// TIA Portal V21 export
// export: Created 2026-11-10T19:21:32.9271764Z, ExportSetting WithDefaults, DisplayName Totally Integrated Automation Portal, DisplayVersion V21 Update 3, DisplayName STEP 7 Professional, DisplayVersion V21 Update 3, DisplayName STEP 7 Safety, DisplayVersion V21, DisplayName Tech WebApplication, DisplayVersion V21, DisplayName WinCC Basic/Comfort/Advanced, DisplayVersion V21 Update 3, DisplayName WinCC Unified, DisplayVersion V21 Update 3
FUNCTION_BLOCK "FB_Lad_pt007"   // FB2, LAD
{ S7_Optimized_Access := 'TRUE' }
VERSION : 0.1
// stored: AutoNumber true, IsIECCheckEnabled false, IsRetainMemResEnabled false, MemoryReserve 100, SetENOAutomatically false, UDAEnableTagReadback false
   VAR_INPUT
      v_req : Bool;
      v_port : PORT;
   END_VAR
   VAR_OUTPUT
      v_ndr : Bool;
      v_dtr : Bool;
      v_dsr : Bool;
      v_rts : Bool;
      v_cts : Bool;
      v_dcd : Bool;
      v_ring : Bool;
      v_error : Bool;
      v_status : Word;
   END_VAR
   VAR
      inst { S7_SetPoint := 'True'} : Signal_Get;
   END_VAR
BEGIN

REGION Network 1: SGN_GET - Query RS-232 signals
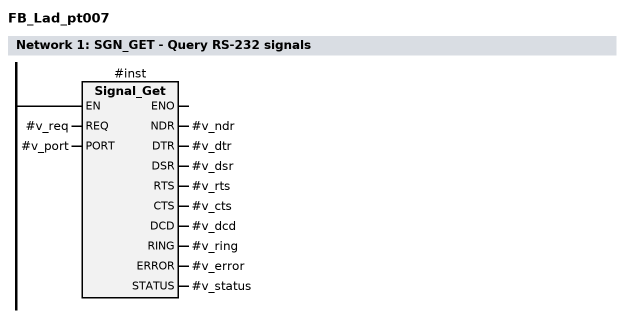
   RUNG wire#powerrail
      #inst.Signal_Get(REQ := #v_req, PORT := #v_port, NDR => #v_ndr, DTR => #v_dtr, DSR => #v_dsr, RTS => #v_rts, CTS => #v_cts, DCD => #v_dcd, RING => #v_ring, ERROR => #v_error, STATUS => #v_status)
   END_RUNG
   // the same network as SCL:
   #inst(REQ := #v_req,   // Signal_Get
         PORT := #v_port,
         NDR => #v_ndr,
         DTR => #v_dtr,
         DSR => #v_dsr,
         RTS => #v_rts,
         CTS => #v_cts,
         DCD => #v_dcd,
         RING => #v_ring,
         ERROR => #v_error,
         STATUS => #v_status);
END_REGION
END_FUNCTION_BLOCK
